// TIA Portal V15.1 export
// export: Created 2000-01-01T00:00:00.0000000Z, ExportSetting None
FUNCTION "FC_Rung" : Void   // FC42, LAD
{ S7_Optimized_Access := 'TRUE' }
   VAR_INPUT
      Local : Int;
   END_VAR
BEGIN

REGION Network 1
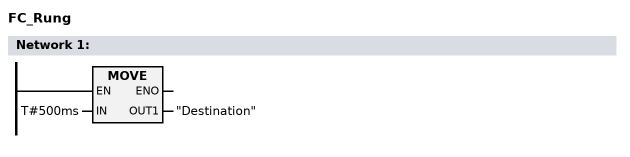
   RUNG wire#powerrail
      Move(in := T#500ms, out1 => "Destination")
   END_RUNG
   // the same network as SCL:
   "Destination" := T#500ms;
END_REGION
END_FUNCTION
